// TIA Portal V14 SP1 export
// export: Created 2000-01-01T00:00:00.0000000Z, ExportSetting None
FUNCTION "FC_Rung" : Void   // FC42, LAD
{ S7_Optimized_Access := 'TRUE' }
   VAR_INPUT
      Local : Int;
   END_VAR
BEGIN

REGION Network 1
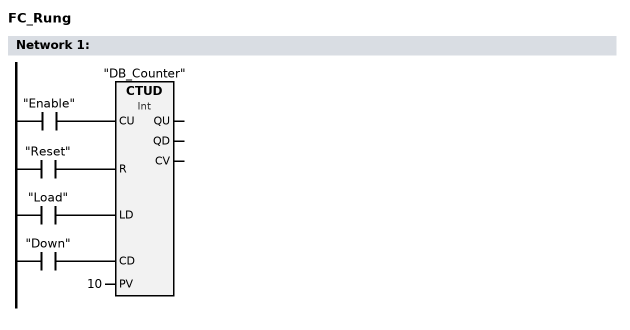
   RUNG wire#powerrail
      Contact( "Enable" )
      { S7_Templates := "value_type := Int" } "DB_Counter".CTUD(r := wire#w1, ld := wire#w2, cd := wire#w3, pv := 10, qd =>, cv =>)
   END_RUNG
   RUNG wire#powerrail
      Contact( "Reset" )
   END_RUNG wire#w1
   RUNG wire#powerrail
      Contact( "Load" )
   END_RUNG wire#w2
   RUNG wire#powerrail
      Contact( "Down" )
   END_RUNG wire#w3
   // the same network as SCL:
   "DB_Counter".CTUD(CU := "Enable", R := "Reset", LD := "Load", CD := "Down", PV := 10);
END_REGION
END_FUNCTION
